Fanuc KAREL source: KT00462.KL

PROGRAM KT00462
%NOLOCKGROUP
VAR
  P1: XYZWPR
  P2: JOINTPOS
  OUT: BOOLEAN
BEGIN
  P1.X = 1.0
  OUT = P1 >= P2
END KT00462
